Staubli VAL3: start.pgx

program start()
begin
  resetMotion(jDepart)
  bInit_repere = false
  taskCreate "IHM",10,IHM()
  call exercice6()
end
